(* IEC 61131-3 sources: trust-platform/examples/rust_service/src/generated, 1 file *)

(* ---- services.st ---- *)
(* GENERATED by trust-runtime from trust.toml - do not edit *)
VAR_GLOBAL
    price_heartbeat : UDINT;
END_VAR
